FUNCTION_BLOCK StationMode (* Basic Function Block Type *)
  (* Standard: 61499-2 *)
  (* Version 0.0, 11/16/2026, Sandeep Patil, Flexbridge AB, Template *)
  PACKAGE Flexbridge.FestoMPS400;
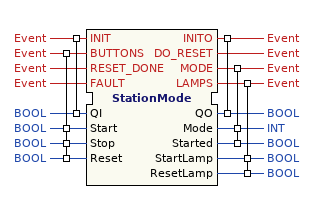
  EVENT_INPUT
    INIT WITH QI; (* Initialisation request *)
    BUTTONS WITH Start, Stop, Reset; (* Console buttons changed *)
    RESET_DONE; (* The station's reset sequence has finished *)
    FAULT; (* The station's sequence stopped on a device fault *)
  END_EVENT
  EVENT_OUTPUT
    INITO WITH QO; (* Initialisation confirm *)
    DO_RESET; (* Start the station's reset sequence *)
    MODE WITH Mode, Started; (* Station mode changed *)
    LAMPS WITH StartLamp, ResetLamp; (* Lamp states for the console *)
  END_EVENT
  VAR_INPUT
    QI : BOOL; (* Input event qualifier *)
    Start : BOOL; (* START button pressed *)
    Stop : BOOL; (* STOP button pressed (already inverted: TRUE while pressed) *)
    Reset : BOOL; (* RESET button pressed *)
  END_VAR
  VAR_OUTPUT
    QO : BOOL; (* Output event qualifier *)
    Mode : INT; (* Station mode: 0 = wait for RESET, 1 = resetting, 2 = wait for START, 3 = started *)
    Started : BOOL; (* TRUE while the station is started and accepts requests *)
    StartLamp : BOOL; (* START lamp *)
    ResetLamp : BOOL; (* RESET lamp *)
  END_VAR
  VAR
    PrevStart : BOOL; (* Start at the last BUTTONS event *)
    PrevStop : BOOL; (* Stop at the last BUTTONS event *)
    PrevReset : BOOL; (* Reset at the last BUTTONS event *)
    StartPressed : BOOL; (* Rising edge of Start *)
    StopPressed : BOOL; (* Rising edge of Stop *)
    ResetReleased : BOOL; (* Falling edge of Reset *)
  END_VAR
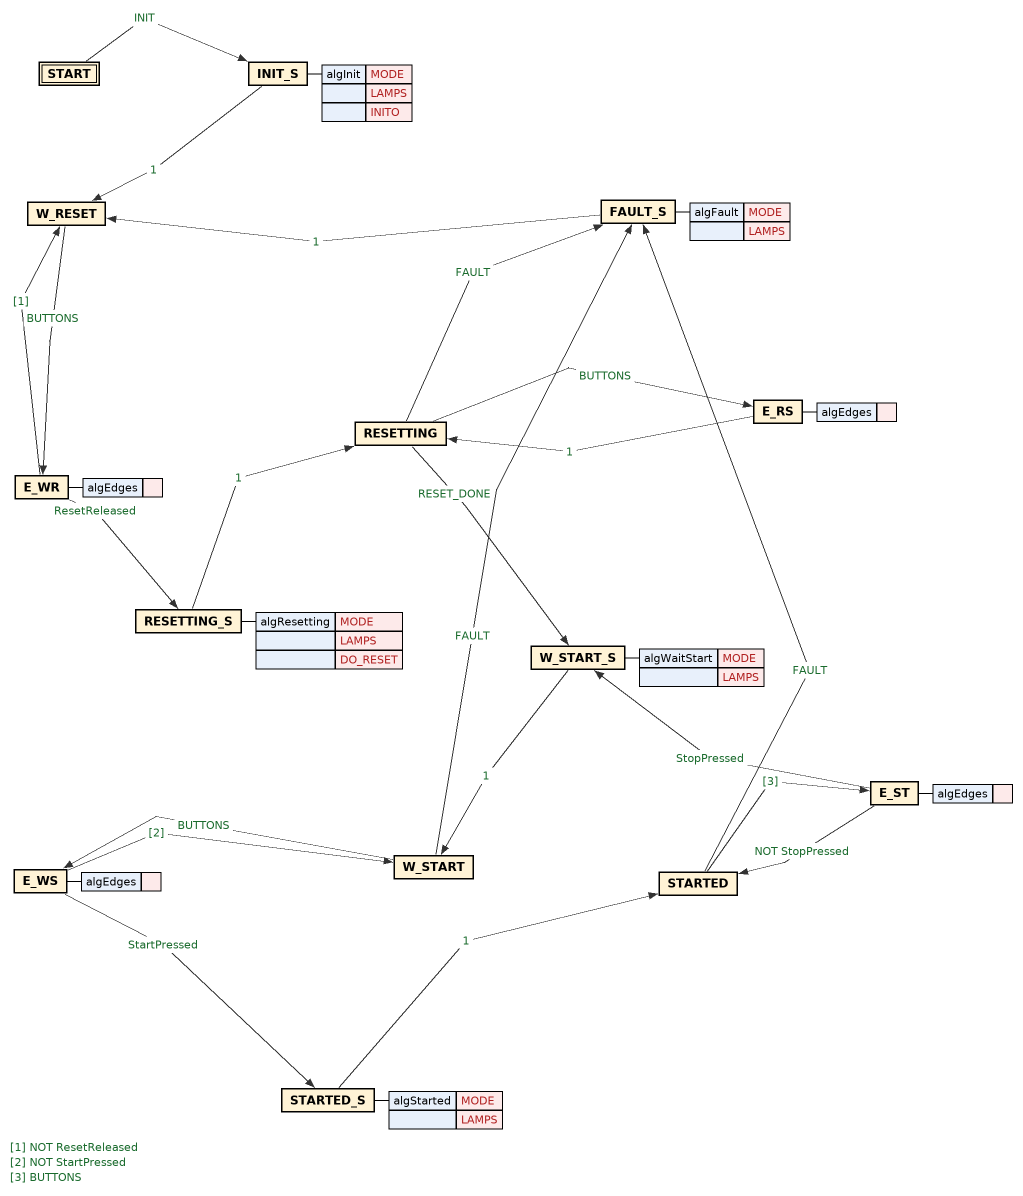
  EC_STATES
    START; (* Initial state *)
    INIT_S : algInit -> MODE, -> LAMPS, -> INITO;
    W_RESET; (* Mode 0: wait for RESET *)
    E_WR : algEdges;
    RESETTING_S : algResetting -> MODE, -> LAMPS, -> DO_RESET;
    RESETTING; (* Mode 1: reset sequence running *)
    E_RS : algEdges;
    W_START_S : algWaitStart -> MODE, -> LAMPS;
    W_START; (* Mode 2: wait for START *)
    E_WS : algEdges;
    STARTED_S : algStarted -> MODE, -> LAMPS;
    STARTED; (* Mode 3: started *)
    E_ST : algEdges;
    FAULT_S : algFault -> MODE, -> LAMPS;
  END_STATES
  EC_TRANSITIONS
    START TO INIT_S := INIT;
    INIT_S TO W_RESET := 1;
    W_RESET TO E_WR := BUTTONS;
    E_WR TO RESETTING_S := ResetReleased;
    E_WR TO W_RESET := NOT ResetReleased;
    RESETTING_S TO RESETTING := 1;
    RESETTING TO W_START_S := RESET_DONE;
    RESETTING TO FAULT_S := FAULT;
    RESETTING TO E_RS := BUTTONS;
    E_RS TO RESETTING := 1;
    W_START_S TO W_START := 1;
    W_START TO E_WS := BUTTONS;
    E_WS TO STARTED_S := StartPressed;
    E_WS TO W_START := NOT StartPressed;
    W_START TO FAULT_S := FAULT;
    STARTED_S TO STARTED := 1;
    STARTED TO E_ST := BUTTONS;
    E_ST TO W_START_S := StopPressed;
    E_ST TO STARTED := NOT StopPressed;
    STARTED TO FAULT_S := FAULT;
    FAULT_S TO W_RESET := 1;
  END_TRANSITIONS
  ALGORITHM algInit IN ST: (* Wait for RESET: RESET lamp on *)
QO := QI;
PrevStart := FALSE; PrevStop := FALSE; PrevReset := FALSE;
StartPressed := FALSE; StopPressed := FALSE; ResetReleased := FALSE;
Mode := 0; Started := FALSE;
StartLamp := FALSE; ResetLamp := TRUE;
  END_ALGORITHM
  ALGORITHM algEdges IN ST: (* Edges of the buttons since the last BUTTONS event *)
StartPressed := Start AND NOT PrevStart;
StopPressed := Stop AND NOT PrevStop;
ResetReleased := PrevReset AND NOT Reset;
PrevStart := Start; PrevStop := Stop; PrevReset := Reset;
  END_ALGORITHM
  ALGORITHM algResetting IN ST: (* Reset sequence running: RESET lamp stays on *)
Mode := 1; Started := FALSE;
StartLamp := FALSE; ResetLamp := TRUE;
  END_ALGORITHM
  ALGORITHM algWaitStart IN ST: (* Wait for START: START lamp on *)
Mode := 2; Started := FALSE;
StartLamp := TRUE; ResetLamp := FALSE;
  END_ALGORITHM
  ALGORITHM algStarted IN ST: (* Started: lamps off *)
Mode := 3; Started := TRUE;
StartLamp := FALSE; ResetLamp := FALSE;
  END_ALGORITHM
  ALGORITHM algFault IN ST: (* Device fault: back to wait for RESET *)
Mode := 0; Started := FALSE;
StartLamp := FALSE; ResetLamp := TRUE;
  END_ALGORITHM
END_FUNCTION_BLOCK
